// Function block for calculating the product of two values
FUNCTION_BLOCK FB_Prod
VAR_INPUT
	var1: UINT;    // variable 1
	var2: UINT;    // variable 2
END_VAR
VAR_OUTPUT
	result : UINT; // result
END_VAR

// Calculation of the product of two values
result := var1 * var2;

END_FUNCTION_BLOCK

(* stored: Version 1.1.0.1, ProductVersion 3.1.4026.18
   POU FB_Prod: Id {00a1861b-3b8e-4d3a-95d3-7f3b2848d738}, SpecialFunc None *)
